Fanuc KAREL source: KO00113.KL

PROGRAM KO00113
%NOLOCKGROUP
VAR
  A: ARRAY[2] OF BYTE
  B: INTEGER
  OUT: INTEGER
BEGIN
  A[1] = 1
  B = 2
  OUT = ATAN2(A[1], B)
END KO00113
